// TIA Portal V20 export
// export: Created 2026-10-12T05:42:35.8894891Z, ExportSetting WithDefaults, DisplayName Totally Integrated Automation Portal, DisplayVersion V20, DisplayName TIA Portal Openness, DisplayVersion V20, DisplayName TIA Portal Teamcenter Gateway, DisplayVersion V20, DisplayName TIA Portal Version Control Interface, DisplayVersion V20, DisplayName SINAMICS Startdrive Advanced, DisplayVersion V20 SP1 Update 2, DisplayName SINAMICS Startdrive G110M, G120, G120C, G120D, G120P, G115D, DisplayVersion V20 SP1 Update 2, DisplayName SINAMICS Startdrive G130, G150, S120, S150, SINAMICS MV, G220, S200, S210, DisplayVersion V20 SP1 Update 2, DisplayName STEP 7 Professional, DisplayVersion V20, DisplayName STEP 7 Safety, DisplayVersion V20, DisplayName WinCC Basic/Comfort/Advanced, DisplayVersion V20, DisplayName WinCC Professional, DisplayVersion V20, DisplayName WinCC Unified, DisplayVersion V20
DATA_BLOCK "GDB_PressDemoIO"   // DB19
{ S7_Optimized_Access := 'TRUE' }
VERSION : 0.1
// Demo logical I/O boundary. Bind these symbols to the commissioned hardware
//  driver when a bench is available; feedback is never synthesized here.
// stored: AutoNumber true, DBAccessibleFromOPCUA true, DBAccessibleFromWebserver true, IsOnlyStoredInLoadMemory false, IsRetainMemResEnabled false, IsWriteProtectedInAS false, MemoryReserve 100
   VAR
      PartPresent : Bool;
      PartQuality : Bool;
      AirPressureOk : Bool;
      TwoHandHeld : Bool;
      StartPulse : Bool;
      RamExtended : Bool;
      RamRetracted : Bool;
      DoorClosed : Bool;
      DoorOpen : Bool;
      SlideInside : Bool;
      SlideOutside : Bool;
      RamExtend : Bool;
      RamRetract : Bool;
      DoorClose : Bool;
      DoorRelease : Bool;
      SlideExtend : Bool;
      SlideRetract : Bool;
   END_VAR
BEGIN
END_DATA_BLOCK
